Fanuc KAREL source: KA00099.KL

PROGRAM KA00099
%NOLOCKGROUP
VAR
  SRC: VECTOR
  DST: BOOLEAN
BEGIN
  SRC.X = 1.0
  DST = SRC
END KA00099
